Fanuc KAREL source: kt00903.KL

-- PROVISIONAL review KL for V940-1; original PC SHA256 cee69815df799477cb01088d7e08fcb6a85bef8fdce665fec099540c33b0035c
-- Incomplete behavior may be omitted. Consult companion uncertainty JSON. Do not deploy.
PROGRAM KT00903
%NOLOCKGROUP
BEGIN
  -- V9_ZERO_TABLE_METADATA_HINT layout=0002_ascii; no indexed target words; source/name/runtime held
  -- UNRESOLVED_PC offsets 5-28; opcodes 27,22,1C,31,4A
  -- UNRESOLVED_PC offsets 33-37; opcodes 7F
END KT00903
